Fanuc KAREL source: KT00844.KL

PROGRAM KT00844
%NOLOCKGROUP
VAR
  I1: INTEGER
  I2: INTEGER
  OUT: INTEGER
BEGIN
  I1 = 2
  I2 = 3
  I1 = 2
  I2 = 3
  OUT = TAN(I1)
END KT00844
